// Mitsubishi GX Works2 project: Task3_Ex_1   PLC: FX3G

PROGRAM MAIN
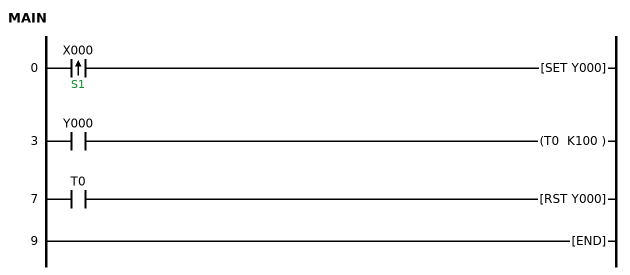
0     LDP     X000  ; S1
      SET     Y000
3     LD      Y000
      OUT     T0 K100
7     LD      T0
      RST     Y000
9     END
END_PROGRAM
